// Mitsubishi GX Works2 project: Control-Robot -Gantry   PLC: Q06UDEH

// task Task_01 (event TRUE, interval 0, priority 31): POU_01
// task PLC_VIS_Ready (event TRUE, interval 0, priority 31): PLC_VIS_Ready
// task Convert_Units (event TRUE, interval 0, priority 31): Convert_Units

PROGRAM Convert_Units
VAR
  Val_Pules : DINT;
  Val_Pules_R : REAL;
  Pules_P : DINT;
  Pules_R : DINT;
  Speed_Conveyor : REAL;
  Circumference : REAL;
  Speed_Conveyor_mm_min : REAL;
END_VAR
VAR CONSTANT
  Const : REAL;
  PPR_R : REAL := 200;  (* Xung\vòng *)
  Diameter_Wheel : REAL := 40.0;  (* D banh xe *)
END_VAR
IF Y0  THEN

    (* === NEAR POINT (K71) === *)
    (* Bit 6 và bit 0 set = Near Point signal *)
    M300 := (D900 = 71);    (* Ax1 Near_Point *)
    M301 := (D901 = 71);    (* Ax2 Near_Point *)
    M302 := (D902 = 71);    (* Ax3 Near_Point *)
    
        (* === LOWER LIMIT (K6) === *)
    (* Bit 2 và bit 1 set = Lower Limit signal *)
    M303 := (D900 = 6);     (* Ax1 Lower_Limit *)
    M304 := (D901 = 6);     (* Ax2 Lower_Limit *)
    M305 := (D902 = 6);     (* Ax3 Lower_Limit *)

    (* === UPPER LIMIT (K5) === *)
    (* Bit 2 và bit 0 set = Upper Limit signal *)
    M306 := (D900 = 5);     (* Ax1 Upper_Limit *)
    M307 := (D901 = 5);     (* Ax2 Upper_Limit *)
    M308 := (D902 = 5);     (* Ax3 Upper_Limit *)

END_IF;

(* Khởi tạo mốc ban đầu ngay khi RUN PLC để chống nhảy số *)
IF SM400 THEN
    DMOV(TRUE, U8\G2, Pules_P);
END_IF;

(* Lấy mẫu tốc độ cao lặp vòng mỗi 100ms *)
IF SM400 THEN
    Y84 := TRUE;
    DMOV(TRUE, U8\G2, D10);
    OUTH_T(TRUE, TC0, 10);

    IF TS0 THEN
        DMOV(TRUE, D10, Pules_R);
        Val_Pules := Pules_R - Pules_P;
        
        Pules_P := Pules_R;             (* Cập nhật mốc mới liên tục *)
        RST(TRUE, TC0);
    END_IF;
END_IF;

(* Tính toán tốc độ *)
IF SM400 THEN
    (* 1. Chỉ ép kiểu duy nhất số xung đo được sang REAL *)
    Val_Pules_R := DINT_TO_REAL(Val_Pules);
    
    (* 2. Tính chu vi bánh xe (mm) *)
    Circumference := 3.14159 * Diameter_Wheel;
       
    (* 3. Tính tốc độ ra mm/phút
       - Do thời gian lấy mẫu là 100ms (0.1s), số xung cần nhân 10.0 để ra số xung/giây.
       - Nhân thêm 60.0 ở cuối để quy đổi từ giây sang phút. *)
    Speed_Conveyor_mm_min := ((Val_Pules_R * 10.0) / PPR_R) * Circumference * 60.0;
END_IF;
END_PROGRAM

PROGRAM PLC_VIS_Ready
VAR CONSTANT
  Const : REAL;
END_VAR
VAR
  Vision_Ready : BOOL;
  PLC_Start : BOOL;
  PLC_Complete : BOOL;
  Vision_Re : BOOL;
  iState : INT;
  diTargetX : DWORD;
  diTargetY : DWORD;
  DONE : BOOL;
  Speed_Conveyor_1 : Speed_Conveyor;
  Tracking_1 : Tracking;
END_VAR
CASE iState OF
    0: (* Bước 0: Chờ sản phẩm và kiểm tra Vision Ready (D3100 = 1) *)
        IF D3100 = 1 THEN
            D3000 := 1; (* PLC Start = 1 *)
            iState := 10;
        END_IF;

    10:

            D3000 := 0; (* Reset PLC Start *)
            D3001 := 1; (* PLC Complete = 1 báo đã nhận dữ liệu *)
            iState := 20;

    20: 
        IF (D3100 = 1) THEN
            D3001 := 0; 
            iState := 0; 
        END_IF;
END_CASE;
END_PROGRAM

PROGRAM POU_01
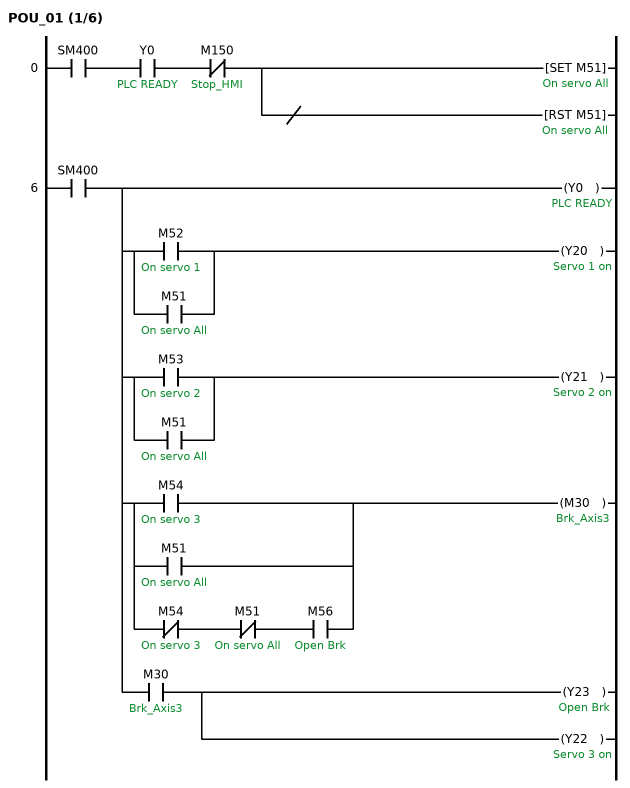
0     LD      SM400
      AND     Y0  ; PLC READY
      ANI     M150  ; Stop_HMI
      SET     M51  ; On servo All
      INV
      RST     M51  ; On servo All
6     LD      SM400
      OUT     Y0  ; PLC READY
      MPS
      LD      M52  ; On servo 1
      OR      M51  ; On servo All
      ANB
      OUT     Y20  ; Servo 1 on
      MRD
      LD      M53  ; On servo 2
      OR      M51  ; On servo All
      ANB
      OUT     Y21  ; Servo 2 on
      MRD
      LD      M54  ; On servo 3
      OR      M51  ; On servo All
      LDI     M54  ; On servo 3
      ANI     M51  ; On servo All
      AND     M56  ; Open Brk
      ORB
      ANB
      OUT     M30  ; Brk_Axis3
      MPP
      AND     M30  ; Brk_Axis3
      OUT     Y23  ; Open Brk
      OUT     Y22  ; Servo 3 on
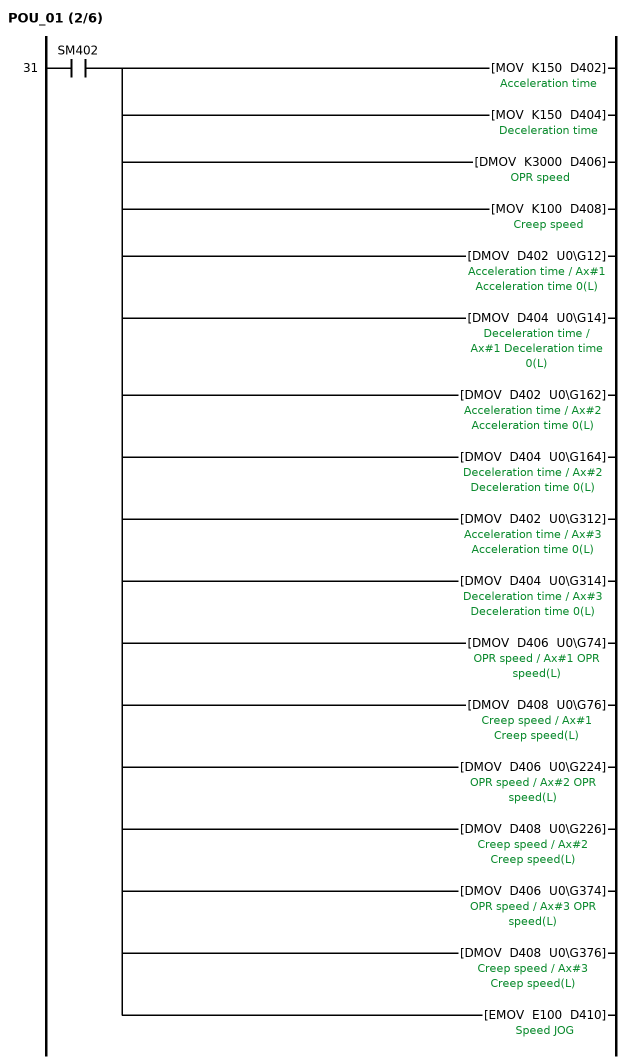
31    LD      SM402
      MOV     K150 D402  ; Acceleration time
      MOV     K150 D404  ; Deceleration time
      DMOV    K3000 D406  ; OPR speed
      MOV     K100 D408  ; Creep speed
      DMOV    D402 U0\G12  ; Ax#1 Acceleration time 0(L)
      DMOV    D404 U0\G14  ; Ax#1 Deceleration time 0(L)
      DMOV    D402 U0\G162  ; Ax#2 Acceleration time 0(L)
      DMOV    D404 U0\G164  ; Ax#2 Deceleration time 0(L)
      DMOV    D402 U0\G312  ; Ax#3 Acceleration time 0(L)
      DMOV    D404 U0\G314  ; Ax#3 Deceleration time 0(L)
      DMOV    D406 U0\G74  ; Ax#1 OPR speed(L)
      DMOV    D408 U0\G76  ; Ax#1 Creep speed(L)
      DMOV    D406 U0\G224  ; Ax#2 OPR speed(L)
      DMOV    D408 U0\G226  ; Ax#2 Creep speed(L)
      DMOV    D406 U0\G374  ; Ax#3 OPR speed(L)
      DMOV    D408 U0\G376  ; Ax#3 Creep speed(L)
      EMOV    E100 D410  ; Speed JOG
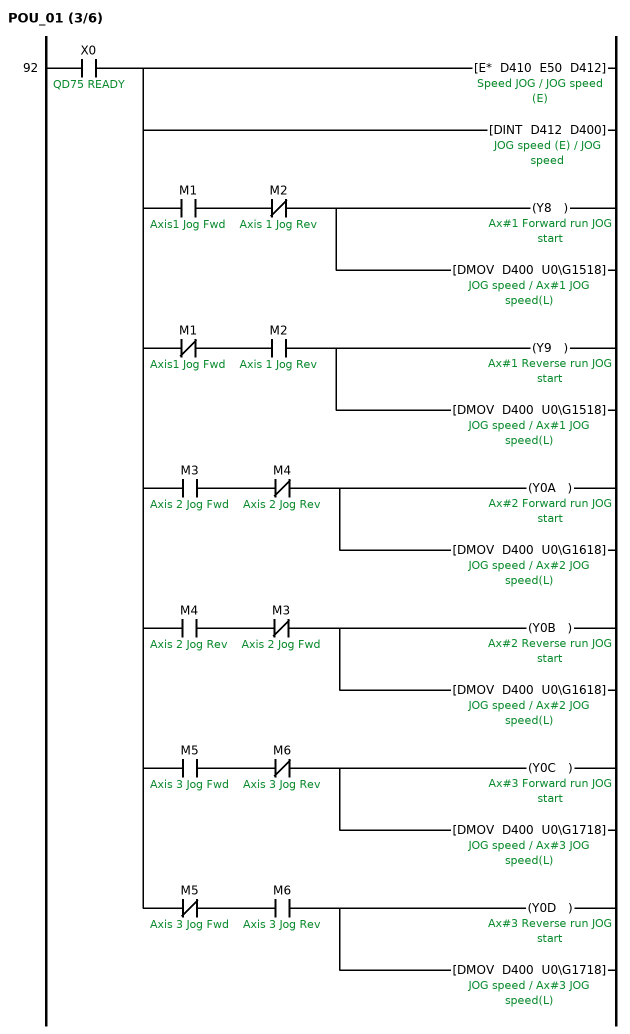
92    LD      X0  ; QD75 READY
      E*      D410 E50 D412  ; JOG speed (E)
      DINT    D412 D400  ; JOG speed
      MPS
      AND     M1  ; Axis1 Jog Fwd
      ANI     M2  ; Axis 1 Jog Rev
      OUT     Y8  ; Ax#1 Forward run JOG start
      DMOV    D400 U0\G1518  ; Ax#1 JOG speed(L)
      MRD
      ANI     M1  ; Axis1 Jog Fwd
      AND     M2  ; Axis 1 Jog Rev
      OUT     Y9  ; Ax#1 Reverse run JOG start
      DMOV    D400 U0\G1518
      MRD
      AND     M3  ; Axis 2 Jog Fwd
      ANI     M4  ; Axis 2 Jog Rev
      OUT     Y0A  ; Ax#2 Forward run JOG start
      DMOV    D400 U0\G1618  ; Ax#2 JOG speed(L)
      MRD
      AND     M4  ; Axis 2 Jog Rev
      ANI     M3  ; Axis 2 Jog Fwd
      OUT     Y0B  ; Ax#2 Reverse run JOG start
      DMOV    D400 U0\G1618
      MRD
      AND     M5  ; Axis 3 Jog Fwd
      ANI     M6  ; Axis 3 Jog Rev
      OUT     Y0C  ; Ax#3 Forward run JOG start
      DMOV    D400 U0\G1718  ; Ax#3 JOG speed(L)
      MPP
      ANI     M5  ; Axis 3 Jog Fwd
      AND     M6  ; Axis 3 Jog Rev
      OUT     Y0D  ; Ax#3 Reverse run JOG start
      DMOV    D400 U0\G1718
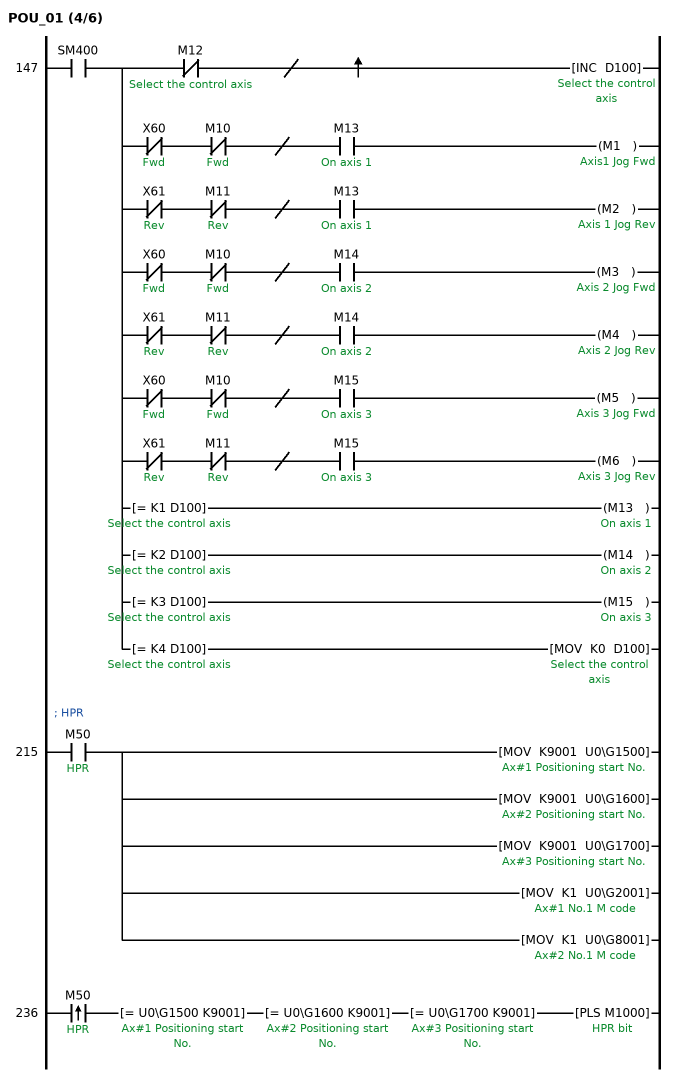
147   LD      SM400
      MPS
      ANI     M12  ; Select the control axis
      INV
      MEP
      INC     D100  ; Select the control axis
      MRD
      ANI     X60  ; Fwd
      ANI     M10  ; Fwd
      INV
      AND     M13  ; On axis 1
      OUT     M1  ; Axis1 Jog Fwd
      MRD
      ANI     X61  ; Rev
      ANI     M11  ; Rev
      INV
      AND     M13  ; On axis 1
      OUT     M2  ; Axis 1 Jog Rev
      MRD
      ANI     X60  ; Fwd
      ANI     M10  ; Fwd
      INV
      AND     M14  ; On axis 2
      OUT     M3  ; Axis 2 Jog Fwd
      MRD
      ANI     X61  ; Rev
      ANI     M11  ; Rev
      INV
      AND     M14  ; On axis 2
      OUT     M4  ; Axis 2 Jog Rev
      MRD
      ANI     X60  ; Fwd
      ANI     M10  ; Fwd
      INV
      AND     M15  ; On axis 3
      OUT     M5  ; Axis 3 Jog Fwd
      MRD
      ANI     X61  ; Rev
      ANI     M11  ; Rev
      INV
      AND     M15  ; On axis 3
      OUT     M6  ; Axis 3 Jog Rev
      MRD
      AND=    K1 D100  ; Select the control axis
      OUT     M13  ; On axis 1
      MRD
      AND=    K2 D100  ; Select the control axis
      OUT     M14  ; On axis 2
      MRD
      AND=    K3 D100  ; Select the control axis
      OUT     M15  ; On axis 3
      MPP
      AND=    K4 D100  ; Select the control axis
      MOV     K0 D100
; HPR
215   LD      M50  ; HPR
      MOV     K9001 U0\G1500  ; Ax#1 Positioning start No.
      MOV     K9001 U0\G1600  ; Ax#2 Positioning start No.
      MOV     K9001 U0\G1700  ; Ax#3 Positioning start No.
      MOV     K1 U0\G2001  ; Ax#1 No.1 M code
      MOV     K1 U0\G8001  ; Ax#2 No.1 M code
236   LDP     M50  ; HPR
      AND=    U0\G1500 K9001  ; Ax#1 Positioning start No.
      AND=    U0\G1600 K9001  ; Ax#2 Positioning start No.
      AND=    U0\G1700 K9001  ; Ax#3 Positioning start No.
      PLS     M1000  ; HPR bit
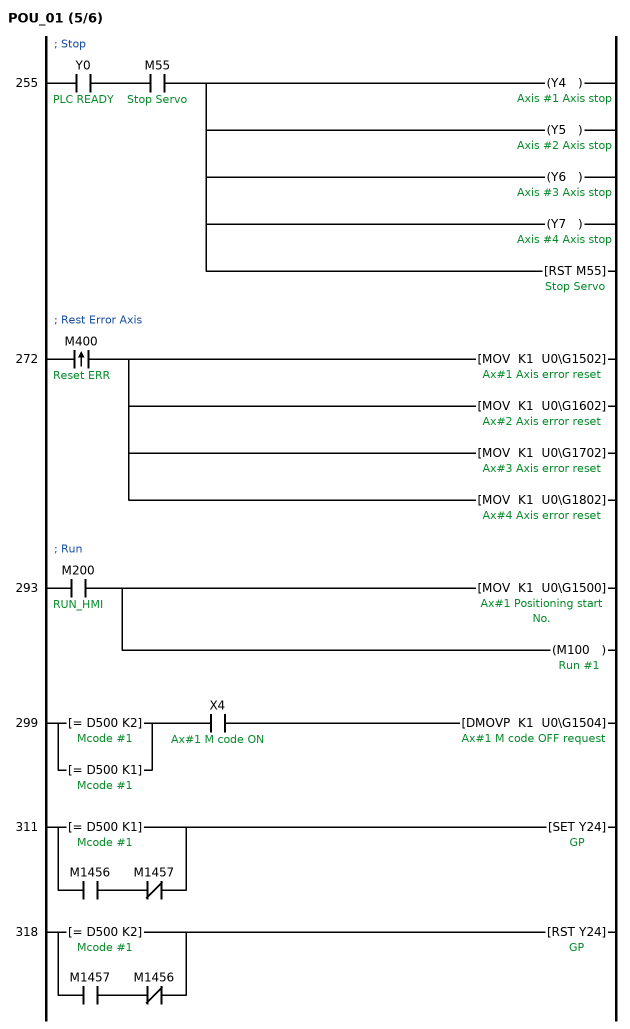
; Stop
255   LD      Y0  ; PLC READY
      AND     M55  ; Stop Servo
      OUT     Y4  ; Axis #1 Axis stop
      OUT     Y5  ; Axis #2 Axis stop
      OUT     Y6  ; Axis #3 Axis stop
      OUT     Y7  ; Axis #4 Axis stop
      RST     M55  ; Stop Servo
; Rest Error Axis
272   LDP     M400  ; Reset ERR
      MOV     K1 U0\G1502  ; Ax#1 Axis error reset
      MOV     K1 U0\G1602  ; Ax#2 Axis error reset
      MOV     K1 U0\G1702  ; Ax#3 Axis error reset
      MOV     K1 U0\G1802  ; Ax#4 Axis error reset
; Run
293   LD      M200  ; RUN_HMI
      MOV     K1 U0\G1500
      OUT     M100  ; Run #1
299   LD=     D500 K2  ; Mcode #1
      OR=     D500 K1  ; Mcode #1
      AND     X4  ; Ax#1 M code ON
      DMOVP   K1 U0\G1504  ; Ax#1 M code OFF request
311   LD=     D500 K1  ; Mcode #1
      LD      M1456
      ANI     M1457
      ORB
      SET     Y24  ; GP
318   LD=     D500 K2  ; Mcode #1
      LD      M1457
      ANI     M1456
      ORB
      RST     Y24  ; GP
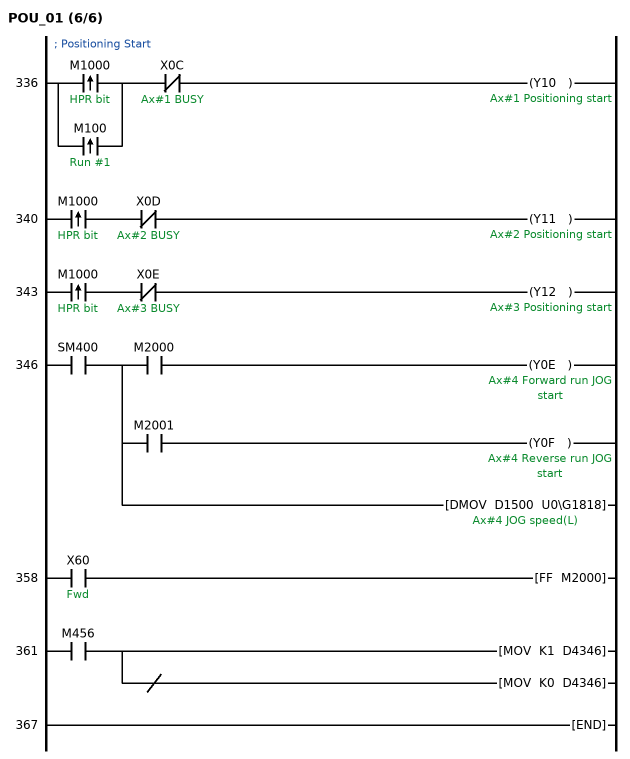
; Positioning Start
336   LDP     M1000  ; HPR bit
      ORP     M100  ; Run #1
      ANI     X0C  ; Ax#1 BUSY
      OUT     Y10  ; Ax#1 Positioning start
340   LDP     M1000  ; HPR bit
      ANI     X0D  ; Ax#2 BUSY
      OUT     Y11  ; Ax#2 Positioning start
343   LDP     M1000  ; HPR bit
      ANI     X0E  ; Ax#3 BUSY
      OUT     Y12  ; Ax#3 Positioning start
346   LD      SM400
      MPS
      AND     M2000
      OUT     Y0E  ; Ax#4 Forward run JOG start
      MRD
      AND     M2001
      OUT     Y0F  ; Ax#4 Reverse run JOG start
      MPP
      DMOV    D1500 U0\G1818  ; Ax#4 JOG speed(L)
358   LD      X60  ; Fwd
      FF      M2000
361   LD      M456
      MOV     K1 D4346
      INV
      MOV     K0 D4346
367   END
END_PROGRAM

FUNCTION_BLOCK Speed_Conveyor
VAR
  Val_Pules : DINT;
  Pules_P : DINT;
  Pules_R : DINT;
  Val_Pules_R : REAL;
  Speed_Conveyor : REAL;
END_VAR
VAR CONSTANT
  Const : REAL;
  PPR_R : REAL := 200;  (* Xung\vòng *)
  Diameter_Wheel : REAL := 40.0;  (* D banh xe *)
END_VAR
VAR
  Circumference : REAL;
END_VAR
VAR_OUTPUT
  Speed_Conveyor_mm_min : REAL;
END_VAR
;
END_FUNCTION_BLOCK

FUNCTION_BLOCK Tracking
VAR
  iState : INT;
  iTracking_State : INT;
  Target_Index : INT;
  Last_Pick_X : DINT;
  Drop_Y_Target : DINT;
  Picked_Count : DINT;
  Enc_Now : DINT;
  Enc_Prev : DINT;
  Enc_Delta : DINT;
  Enc_Cumulative : DINT;
  Enc_Init_Done : BOOL;
  Pulse_Per_MM : REAL;
  Belt_Speed_MM_Min : REAL;
  Scan_Time_Sec : REAL;
  X_Robot : DINT;
  Axis1_Start : BOOL;
  Axis2_Start : BOOL;
  Axis1_Done : BOOL;
  Axis2_Done : BOOL;
  Last_Axis_Done : BOOL;
  Axis_Done_Rise : BOOL;
  X_Min : DINT;
  X_Max : DINT;
  Rev_Threshold : DINT;
  Reverse_Mode : BOOL;
  D3103_Bool : BOOL;
  D3103_Last : BOOL;
  D3103_Rise : BOOL;
  Queue_Enq_Req : BOOL;
  Queue_Deq_Req : BOOL;
  Queue_Deq_Idx : INT;
  Clear_Queue : BOOL;
  Queue_In_X : DINT;
  Queue_In_Y : DINT;
  Queue_In_Enc : DINT;
  Tracker_Active : BOOL;
  Tracker_X_Cam : DINT;
  X_Real : DINT;
  Y_Real : DINT;
  X_Real_0 : DINT;
  Skip_Count : INT;
  Alarm_Q_Full : BOOL;
  Q_Size : INT;
  Q_Count : INT;
  Q_Arr_X : ARRAY [0..19] OF DINT;
  Q_Arr_Y : ARRAY [0..19] OF DINT;
  Q_Arr_Enc : ARRAY [0..19] OF DINT;
  Q_Empty : BOOL;
  Q_Full : BOOL;
  Q_Out_X : DINT;
  Q_Out_Y : DINT;
  Q_Out_Enc : DINT;
  Q_Out_Idx : INT;
  Q_Loop_Idx : INT;
  Q_Shift_Idx : INT;
  Q_Best_Idx : INT;
  Q_Best_Dist : DINT;
  Q_Cur_X : DINT;
  Q_Cur_Dist : DINT;
  Tracker_Accumulated_X : REAL;
  Tracker_Last_Active : BOOL;
  Tracker_Item_X_Real : DINT;
END_VAR
;
END_FUNCTION_BLOCK

// device comments not shown above
Y84  ; CH1 Count enable command
M300  ; Near_Point_#1
M301  ; Near_Point_#2
M302  ; Near_Point_#3
M303  ; Lower_limit_#1
M304  ; Lower_limit_#2
M305  ; Lower_limit_#3
M306  ; Upper_limit_#1
M307  ; Upper_limit_#2
M308  ; Upper_limit_#3
D900  ; I/O_Extemal_#1
D901  ; I/O_Extemal_#2
D902  ; I/O_Extemal_#3
X1  ; Synchronization flag signal
X5  ; Ax#2 M code ON
X6  ; Ax#3 M code ON
X7  ; Ax#4 M code ON
X8  ; Ax#1 Error detection
X9  ; Ax#2 Error detection
X0A  ; Ax#3 Error detection
X0B  ; Ax#4 Error detection
X0F  ; Ax#4 BUSY
X10  ; Ax#1 Start complete
X11  ; Ax#2 Start complete
X12  ; Ax#3 Start complete
X13  ; Ax#4 Start complete
X14  ; Ax#1 Positioning complete
X15  ; Ax#2 Positioning complete
X16  ; Ax#3 Positioning complete
X17  ; Ax#4 Positioning complete
X62  ; On Servo
X63  ; Run
X64  ; S_HPR
X65  ; Stop
X66  ; Select the control axis
X67  ; Run the conveyor
X68  ; Rev conveyor
X69  ; Turn off conveyor
X80  ; Module READY
X81  ; CH1 Cntr val lrg(pt No. 1)
X82  ; CH1 Cntr val coinc(pt No. 1)
X83  ; CH1 Cntr val sml(pt No. 1)
X84  ; CH1 Extrnl prst rqst dtc
X85  ; CH1 Cntr val lrg(pt No. 2)
X86  ; CH1 Cntr val coinc(pt No. 2)
X87  ; CH1 Cntr val sml(pt No. 2)
X88  ; CH2 Cntr val lrg(pt No. 1)
X89  ; CH2 Cntr val coinc(pt No. 1)
X8A  ; CH2 Cntr val sml(pt No. 1)
X8B  ; CH2 Extrnl prst rqst dtc
X8C  ; CH2 Cntr val lrg(pt No. 2)
X8D  ; CH2 Cntr val coinc(pt No. 2)
X8E  ; CH2 Cntr val sml(pt No. 2)
X8F  ; Fuse broken detection flag
Y13  ; Ax#4 Positioning start
Y14  ; Ax#1 Exe prhbtn flag sgnl
Y15  ; Ax#2 Exe prhbtn flag sgnl
Y16  ; Ax#3 Exe prhbtn flag sgnl
Y17  ; Ax#4 Exe prhbtn flag sgnl
Y80  ; CH1 Coinc sgnl No. 1 rst cmd
Y81  ; CH1 Preset command
Y82  ; CH1 Coinc sgnl enbl cmd
Y83  ; CH1 Down count command
Y85  ; CH1 Extrnl prst dtc rst cmd
Y86  ; CH1 Cntr fnctn sel strt cmd
Y87  ; CH1 Coinc sgnl No. 2 rst cmd
Y88  ; CH2 Coinc sgnl No. 1 rst cmd
Y89  ; CH2 Preset command
Y8A  ; CH2 Coinc sgnl enbl cmd
Y8B  ; CH2 Down count command
Y8C  ; CH2 Count enable command
Y8D  ; CH2 Extrnl prst dtc rst cmd
Y8E  ; CH2 Cntr fnctn sel strt cmd
Y8F  ; CH2 Coinc sgnl No. 2 rst cmd
M0  ; Step On
M7  ; Fwd Conveyor belt
M8  ; Run Conveyor belt
M70  ; Fwd conveyor
M71  ; Rev conveyor
M101  ; Run_Tracking
M201  ; RST_HMI
M202  ; Run_Tracking
M309  ; Conveyor_Fwd
M310  ; Conveyor_Rev
M600  ; Rset couter
D0  ; Pos_Axis1
D2  ; Pos_Axis2
D4  ; Pos_Axis3
D502  ; Axis warning No. – Axis 1
D504  ; Axis error No. – Axis 1
D506  ; Axis warning No. – Axis 2
D508  ; Axis error No. – Axis 2
D510  ; Axis warning No. – Axis 3
D512  ; Axis error No. – Axis 3
D600  ; Current feed value – Axis 1
D602  ; Machine feed value – Axis 1
D604  ; Feedrate – Axis 1
D700  ; Current feed value – Axis 2
D702  ; Machine feed value – Axis 2
D704  ; Feedrate – Axis 2
D800  ; Current feed value – Axis 3
D802  ; Machine feed value – Axis 3
D804  ; Feedrate – Axis 3
D2000  ; E_VisionPos_Axis1
D2002  ; E_VisionPos_Axis2
D2004  ; E_VisionPos_Axis3
D2006  ; E_Speed
D3200  ; Pos_Axis1
D3202  ; Pos_Axis2
D3204  ; Pos_Axis3
T0  ; 1
T10  ; Detal t
